FUNCTION_BLOCK logiBUS_QD_PWM_G (* Output service interface function block for 13-bit PWM output with gamma correction for lamps and LEDs (brightness 0..8191 in DWORD) *)
  (* Description: Copyright (c) 2017 fortiss GmbH, HR Agrartechnik GmbH This program and the accompanying materials are made available under the terms of the Eclipse Public License 2.0 which is available at https://www.eclipse.org/legal/epl-2.0/ SPDX-License-Identifier: EPL-2.0 *)
  (* Version 1.0, 2026-11-06, Franz Höpfinger, HR Agrartechnik GmbH, initial version, gamma variant of logiBUS_QD_PWM *)
  PACKAGE logiBUS::io::DQ;
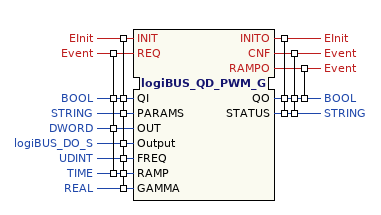
  EVENT_INPUT
    INIT : EInit WITH QI, PARAMS, Output, FREQ, RAMP, GAMMA; (* Service Initialization *)
    REQ WITH QI, OUT, RAMP; (* Service Request *)
  END_EVENT
  EVENT_OUTPUT
    INITO : EInit WITH QO, STATUS; (* Initialization Confirm *)
    CNF WITH QO, STATUS; (* Confirmation of Requested Service *)
    RAMPO WITH QO; (* Ramp finished: OUT reached (immediately after the jump with RAMP = T#0ms) *)
  END_EVENT
  VAR_INPUT
    QI : BOOL; (* Event Input Qualifier *)
    PARAMS : STRING; (* Service Parameters *)
    OUT : DWORD; (* Brightness as the eye sees it (0..8191), converted to the duty cycle with GAMMA, also during the ramp *)
    Output : logiBUS::io::DQ::logiBUS_DO_S := logiBUS_DO::Invalid; (* Identify the Output Output_Q1..Q8 *)
    FREQ : UDINT := 400; (* PWM frequency in Hz, read at INIT. Outputs with the same frequency share an LEDC timer (4 timers, LED blinking uses one). Power stage limits, not checked: APIXON 15 PWR Q1 (BTH50030) max. 100 Hz; BTS7030/BTT6030/BTH6070 for valves 100..200 Hz; Trainer20 without power stage *)
    RAMP : TIME := T#0ms; (* Transition time to the new OUT value (hardware ramp), read at INIT and REQ. T#0ms = jump *)
    GAMMA : REAL := 2.2; (* Gamma of the brightness curve, read at INIT: duty = 8191 * (OUT / 8191)^GAMMA. 1.0 = linear (like logiBUS_QD_PWM), 2.2 = sRGB (default), 2.6 / 2.8 = Espressif examples, often more even on LEDs. Invalid values (<= 0, not finite) run linear like 1.0 *)
  END_VAR
  VAR_OUTPUT
    QO : BOOL; (* Event Output Qualifier *)
    STATUS : STRING; (* Service Status *)
  END_VAR
END_FUNCTION_BLOCK
